FUNCTION_BLOCK SpringMagazineCtrl (* Basic Function Block Type *)
  (* Standard: 61499-2 *)
  (* Version 0.0, 7/2/2026, Template *)
  PACKAGE Main;
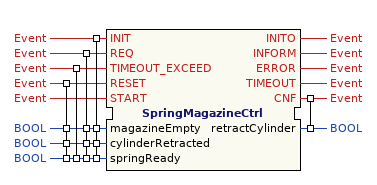
  EVENT_INPUT
    INIT WITH magazineEmpty, cylinderRetracted, springReady; (* Initialization Request *)
    REQ WITH magazineEmpty, cylinderRetracted, springReady; (* Normal Execution Request *)
    TIMEOUT_EXCEED WITH springReady;
    RESET WITH magazineEmpty, cylinderRetracted, springReady;
    START;
  END_EVENT
  EVENT_OUTPUT
    INITO; (* Initialization Confirm *)
    INFORM;
    ERROR;
    TIMEOUT;
    CNF WITH retractCylinder;
  END_EVENT
  VAR_INPUT
    magazineEmpty : BOOL; (* Input event qualifier *)
    cylinderRetracted : BOOL;
    springReady : BOOL;
  END_VAR
  VAR_OUTPUT
    retractCylinder : BOOL;
  END_VAR
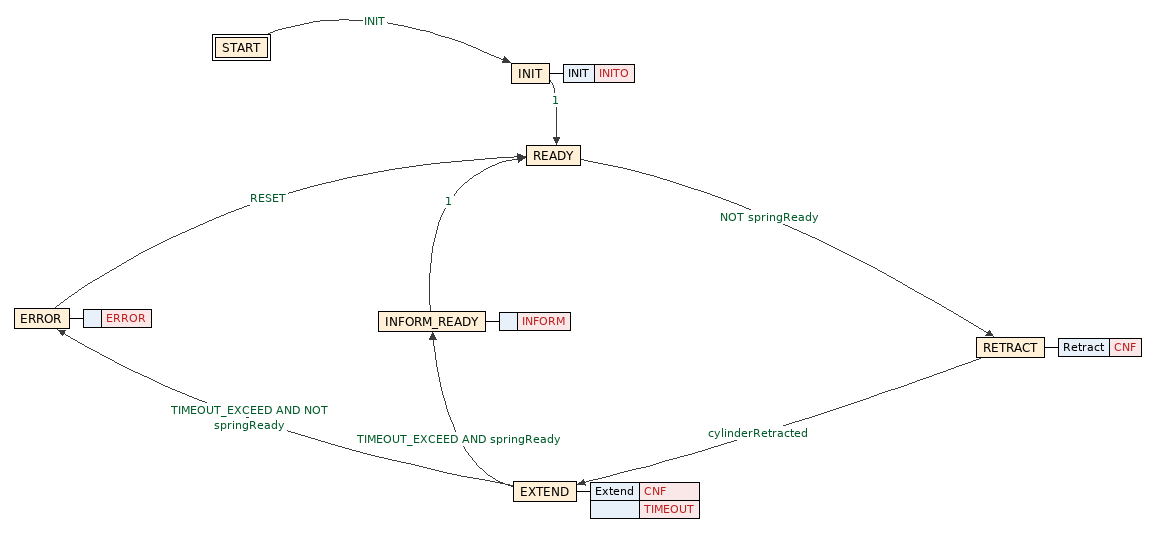
  EC_STATES
    START; (* Initial State *)
    INIT : INIT -> INITO; (* Initialization *)
    READY;
    RETRACT : Retract -> CNF;
    EXTEND : Extend -> CNF, -> TIMEOUT;
    INFORM_READY : -> INFORM;
    ERROR : -> ERROR;
  END_STATES
  EC_TRANSITIONS
    START TO INIT := INIT;
    INIT TO READY := 1;
    READY TO RETRACT := NOT springReady;
    RETRACT TO EXTEND := cylinderRetracted;
    EXTEND TO INFORM_READY := TIMEOUT_EXCEED AND springReady;
    INFORM_READY TO READY := 1;
    EXTEND TO ERROR := TIMEOUT_EXCEED AND NOT springReady;
    ERROR TO READY := RESET;
  END_TRANSITIONS
  ALGORITHM INIT IN ST: (* Initialization algorithm *)
retractCylinder := FALSE;
  END_ALGORITHM
  ALGORITHM REQ IN ST: (* Normally executed algorithm *)
;
  END_ALGORITHM
  ALGORITHM Extend IN ST:
retractCylinder := FALSE;
  END_ALGORITHM
  ALGORITHM Retract IN ST:
retractCylinder := TRUE;
  END_ALGORITHM
END_FUNCTION_BLOCK
